Universal Robots PolyScope program: Prog_Name_That_Is_Very_Long_123.urp

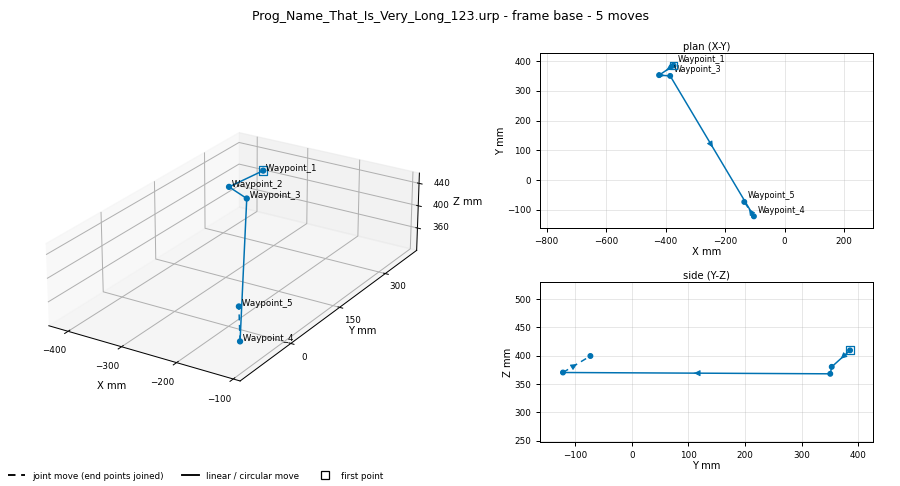
[picture p0: tool path of Prog_Name_That_Is_Very_Long_123.urp in frame base, 5 of 5 moves have a stored position in this frame; points joined in program order, loops and branches not executed]
Program Prog_Name_That_Is_Very_Long_123 (createdIn=3.0.0 lastSavedIn=3.0.0 directory=/programs installation=default)
Robot Program (runOnlyOnce=true motionType=MoveJ speed=1.047198 acceleration=1.396263 useActiveTCP=false)
  'Program generated by VerticalBot Studio for UR5e on 25/10/2026 12:00:00'
  'Using nominal kinematics.'
  'Using Ref. UR5e Base: p[0.000000, 0.000000, 0.000000, 0.000000, 0.000000, 0.000000]'
  'Using TCP Spindle: p[0.010000, 0.000000, 0.120000, 0.000000, 0.261799, 0.000000]'
  Script: set_tcp(p[0.010000, 0.000000, 0.120000, 0.000000, 0.261799, 0.000000])
  Script: movej([-0.523599, -1.745329, 1.570796, -1.396263, -1.570796, 0.349066],1.20000,0.75000,0,0.0000)
  MoveJ speed 42.97 deg/s, acceleration 68.75 deg/s^2 (useActiveTCP=true)
    Waypoint Waypoint_1: TCP in base x=-373.291 y=385.355 z=409.557 mm, rx=-3.0806 ry=-0.2695 rz=-0.4056 rad; joints [-30, -100, 90, -80, -90, 20] deg; flange x=-383.139 y=383.619 z=529.557 mm, rx=3.1296 ry=0.2738 rz=0 rad
  MoveL speed 1000 mm/s, acceleration 1200 mm/s^2 (useActiveTCP=true)
    Waypoint Waypoint_2: motionParameters(blendRadius=0.01); TCP in base x=-421.76 y=353.029 z=380.392 mm, rx=3.0485 ry=0.4964 rz=0.4546 rad; joints [-22, -96, 90, -80, -90, 20] deg; flange x=-436.419 y=356.529 z=499.861 mm, rx=3.0422 ry=0.4818 rz=0.0521 rad
    Waypoint Waypoint_3: motionParameters(blendRadius=0.001); TCP in base x=-384.494 y=350.433 z=368.074 mm, rx=3.0368 ry=0.3896 rz=0.4617 rad; joints [-26, -100, 95, -80, -90, 20] deg; flange x=-400.038 y=356.674 z=487.319 mm, rx=3.0404 ry=0.3733 rz=0.0607 rad
  Halt
  Wait Sleep waitTime=1.5
  Popup Message (haltProgram=false message=Say "hi" to the operator)
  'A long comment line that exceeds the usual controller limits for comments by far, really'
  Set DigitalOutput pin=digital_out[12]; digitalValue=0
  Set DigitalOutput pin=OUT_A; digitalValue=1
  Wait DigitalInput pin=digital_in[get_standard_digital_in(4)]; digitalValue=0
  Wait DigitalInput pin=IN_B; digitalValue=1
  Call Program_With_A_Long_Name_ABCDEFGHIJ
  'Using Ref. Frame 12: p[0.250000, 0.300000, -0.010000, 0.000000, 0.000000, 1.570796]'
  'Using TCP Tool 7: p[0.010000, 0.000000, 0.120000, 0.000000, 0.261799, 0.000000]'
  Script: set_tcp(p[0.010000, 0.000000, 0.120000, 0.000000, 0.261799, 0.000000])
  MoveL speed 1000 mm/s, acceleration 1200 mm/s^2 (useActiveTCP=true)
    Waypoint Waypoint_4: motionParameters(blendRadius=0.001); TCP in base x=-103.029 y=-121.76 z=370.392 mm, rx=-1.7127 ry=-2.3789 rz=-0.3257 rad; joints [-22, -96, 90, -80, -90, 20] deg; flange x=-106.529 y=-136.419 z=489.861 mm, rx=1.8342 ry=2.5246 rz=0.1048 rad
  Script: movej([-0.523599, -1.745329, 1.570796, -1.396263, -1.570796, 0.349066],1.74533,0.52360,0,0.0000)
  MoveJ speed 30.02 deg/s, acceleration 99.98 deg/s^2 (useActiveTCP=true)
    Waypoint Waypoint_5: TCP in base x=-135.355 y=-73.291 z=399.557 mm, rx=-1.8839 ry=-2.2451 rz=-0.248 rad; joints [-30, -100, 90, -80, -90, 20] deg; flange x=-133.619 y=-83.139 z=519.557 mm, rx=2.0194 ry=2.4066 rz=0 rad
SubProgram  [hidden by the author, left out]
SubProgram Program_With_A_Long_Name_ABCDEFGHIJ [hidden by the author, left out]
